Fanuc KAREL source: ko00066.KL

-- PROVISIONAL review KL for V770-1; original PC SHA256 5ac349706edea123a88089b1974842fb202284f9a27b97910d2a679b592e4645
-- Incomplete behavior may be omitted. Consult companion uncertainty JSON. Do not deploy.
PROGRAM KO00066
%NOLOCKGROUP
BEGIN
  -- UNRESOLVED_PC offsets 5-12; opcodes 9D,23
  -- UNRESOLVED_PC offsets 17-63; opcodes 27,22,1C,22,1C,22,31,7E,4A
  -- UNRESOLVED_PC offsets 68-72; opcodes 7F
END KO00066
